Staubli VAL3: applyLib.pgx

public program applyLib()
begin
  savedata:bLibApplied=!savedata:bLibApplied
  savedata:libSave()
  delay(0.5)

end
